// TIA Portal V21 export
// export: Created 2026-11-10T07:35:02.6954762Z, ExportSetting WithDefaults, DisplayName Totally Integrated Automation Portal, DisplayVersion V21 Update 3, DisplayName STEP 7 Professional, DisplayVersion V21 Update 3, DisplayName STEP 7 Safety, DisplayVersion V21, DisplayName Tech WebApplication, DisplayVersion V21, DisplayName WinCC Basic/Comfort/Advanced, DisplayVersion V21 Update 3, DisplayName WinCC Unified, DisplayVersion V21 Update 3
FUNCTION_BLOCK "FB_Lad_ex015"   // FB12, LAD
{ S7_Optimized_Access := 'TRUE' }
VERSION : 0.1
// stored: AutoNumber true, IsIECCheckEnabled false, IsRetainMemResEnabled false, MemoryReserve 100, SetENOAutomatically false, UDAEnableTagReadback false
   VAR_INPUT
      v_in : String;
   END_VAR
   VAR_OUTPUT
      v_out : String;
   END_VAR
BEGIN

REGION Network 1: S_MOVE - Move character string
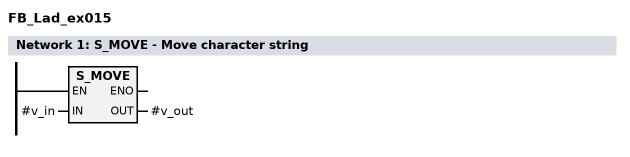
   RUNG wire#powerrail
      S_Move(in := #v_in, out => #v_out)
   END_RUNG
   // the same network as SCL:
   #v_out := #v_in;
END_REGION
END_FUNCTION_BLOCK
